// TIA Portal V21 export
// export: Created 2026-10-24T16:30:26.0512449Z, ExportSetting WithDefaults, DisplayName Totally Integrated Automation Portal, DisplayVersion V21 Update 1, DisplayName SINAMICS Startdrive Advanced, DisplayVersion V21 HF2, DisplayName SINAMICS Startdrive G110M, G120, G120C, G120D, G120P, G115D, DisplayVersion V21 HF2, DisplayName SINAMICS Startdrive G130, G150, S120, S150, G200, G220, S200, S210, S220, Innomotics MVD, DisplayVersion V21 HF2, DisplayName STEP 7 Professional, DisplayVersion V21 Update 1, DisplayName STEP 7 Safety, DisplayVersion V21, DisplayName Tech WebApplication, DisplayVersion V21, DisplayName WinCC Basic/Comfort/Advanced, DisplayVersion V21 Update 1, DisplayName WinCC Unified, DisplayVersion V21 Update 1
TYPE "UDT_V4_Point"
// stored: IsFailsafeCompliant false
   STRUCT
      X : Real;   // Horizontal position
      Y : Real;   // Vertical position
   END_STRUCT;
END_TYPE
